FUNCTION_BLOCK fbShutterCmdSourceSwitch 
VAR_INPUT
    OpenSwitchState : stSwitchState;
    CloseSwitchState : stSwitchState;
    ShutterStateType : eShutterStateType;
END_VAR
VAR_OUTPUT
	Cmd : stShutterCommand;
	NewCmd : BOOL;
END_VAR
VAR
    UpLongClickPosition : stShutterPosition := (Height := 50, Angle := 100);
    DownLongClickPosition : stShutterPosition := (Height := 0, Angle := 100);
END_VAR


// Default outputs every cycle
Cmd.CommandType := eShutterCommandType.NONE;
Cmd.Position.Height := 0;
Cmd.Position.Angle := 0;
NewCmd := FALSE;

// If shutter is moving, any button event means STOP
IF (ShutterStateType <> eShutterStateType.IDLE)
   AND (
        (OpenSwitchState.StateType <> eSwitchStateType.IDLE)
        OR
        (CloseSwitchState.StateType <> eSwitchStateType.IDLE)
   ) THEN
    Cmd.CommandType := eShutterCommandType.STOP;
    NewCmd := TRUE;

// OPEN: double click UP
ELSIF (OpenSwitchState.StateType = eSwitchStateType.MULTI_CLICK)
   AND (OpenSwitchState.PressCount = 2) THEN
    Cmd.CommandType := eShutterCommandType.OPEN;
    NewCmd := TRUE;

// CLOSE: double click DOWN
ELSIF (CloseSwitchState.StateType = eSwitchStateType.MULTI_CLICK)
   AND (CloseSwitchState.PressCount = 2) THEN
    Cmd.CommandType := eShutterCommandType.CLOSE;
    NewCmd := TRUE;

// STEP_OPEN: short click UP
ELSIF OpenSwitchState.StateType = eSwitchStateType.SHORT_CLICK THEN
    Cmd.CommandType := eShutterCommandType.STEP_OPEN;
    NewCmd := TRUE;

// STEP_CLOSE: short click DOWN
ELSIF CloseSwitchState.StateType = eSwitchStateType.SHORT_CLICK THEN
    Cmd.CommandType := eShutterCommandType.STEP_CLOSE;
    NewCmd := TRUE;

// MOVE_TO_POSITION: long click UP
ELSIF (OpenSwitchState.StateType = eSwitchStateType.LONG_CLICK) THEN
    Cmd.CommandType := eShutterCommandType.MOVE_TO_POSITION;
    Cmd.Position := UpLongClickPosition;
    NewCmd := TRUE;
	// MOVE_TO_POSITION: long click DOWN
ELSIF (CloseSwitchState.StateType = eSwitchStateType.LONG_CLICK) THEN
    Cmd.CommandType := eShutterCommandType.MOVE_TO_POSITION;
    Cmd.Position := DownLongClickPosition;
    NewCmd := TRUE;
END_IF

END_FUNCTION_BLOCK

(* stored: Version 1.1.0.1
   POU fbShutterCmdSourceSwitch: Id {6425a77e-86b3-44e6-82a6-6f2235e7d8cd}, SpecialFunc None *)
